{attribute 'qualified_only'}
{attribute 'strict'}
{attribute 'to_string'}
TYPE E_LogRecordFlag:
(
	// The zero value for the enum. Should not be used for comparisons.
	// Instead use bitwise "and" with the appropriate mask as shown above.
	LOG_RECORD_FLAGS_DO_NOT_USE := 0,
	// Bits 0-7 are used for trace flags.
	LOG_RECORD_FLAGS_TRACE_FLAGS_MASK := 255 //0x000000FF;
) UDINT;
END_TYPE
//  LOG_RECORD_FLAGS_TRACE_FLAGS_MASK = '255 '

(* stored: Version 1.1.0.1
   EnumerationTextList E_LogRecordFlag: Id {f9f2013c-0001-4579-8868-ee61015442e4} *)
